DATA_BLOCK "ControlNodes"
{ S7_Optimized_Access := 'TRUE' }
VERSION : 0.1
NON_RETAIN
STRUCT
    sequence : "LAF_typeSequence";
    jobs : "LAF_typeJobs";
    cylFC2400VisualCalibrationFeed : "LBC_TwoWayActuatorControlNodes";
    sensorFC2400VisualCalibrationReady : "LBC_DigitalSignalControlNodes";
END_STRUCT;
BEGIN
END_DATA_BLOCK
